// TIA Portal V20 export
VAR_GLOBAL   // PLC tag table "standard"
   SIMULACE AT %M2.0 : Bool;
   LOG_0 AT %M2.1 : Bool;
   LOG_1 AT %M2.2 : Bool;
   SMAZ_ME_0 AT %M2.3 : Bool;
   SMAZ_ME_1 AT %M2.4 : Bool;
   AUTOMAT AT %M2.5 : Bool;
   MANUAL AT %M2.6 : Bool;
   INICIALIZACE_OK AT %M3.3 : Bool;
   INICIALIZACE AT %M3.4 : Bool;
   INICIALIZACE_RUN AT %M3.5 : Bool;
   LINE_READY_START AT %M3.6 : Bool;
   alrm_global AT %M3.2 : Bool;
   wrong_global AT %M3.7 : Bool;
   alrm_op_0 AT %M4.0 : Bool;
   wrong_op_0 AT %M4.1 : Bool;
   alrm_op_1 AT %M4.2 : Bool;
   wrong_op_1 AT %M4.3 : Bool;
   I_i AT %MW6 : Int;
   "I_i(1)" AT %MW8 : Int;
   adresace AT %MW12 : Int;
   byte_smazat AT %MB5 : Byte;
   inicializace_block AT %M4.4 : Bool;
   s2_hsc_hrana AT %M4.5 : Bool;
   hodnota_volitelna AT %MB14 : Byte;
   Clock_Byte AT %MB0 : Byte;
   Clock_10Hz AT %M0.0 : Bool;
   Clock_5Hz AT %M0.1 : Bool;
   "Clock_2.5Hz" AT %M0.2 : Bool;
   Clock_2Hz AT %M0.3 : Bool;
   "Clock_1.25Hz" AT %M0.4 : Bool;
   Clock_1Hz AT %M0.5 : Bool;
   "Clock_0.625Hz" AT %M0.6 : Bool;
   "Clock_0.5Hz" AT %M0.7 : Bool;
   System_Byte AT %MB1 : Byte;
   FirstScan AT %M1.0 : Bool;
   DiagStatusUpdate AT %M1.1 : Bool;
   AlwaysTRUE AT %M1.2 : Bool;
   AlwaysFALSE AT %M1.3 : Bool;
   INICIALIZACE_REPEAT AT %M4.6 : Bool;
   AUT_MAN_HMI AT %M4.7 : Bool;   // POUŽÍVÁNO PRO PANELOUVOU VOLBU
   volny_pristup_2 AT %M10.0 : Bool;
   alrm_op_2 AT %M11.3 : Bool;
   wrong_op_2 AT %M11.4 : Bool;
   alrm_op_3 AT %M11.5 : Bool;
   wrong_op_3 AT %M11.6 : Bool;
   alrm_op_4 AT %M11.7 : Bool;
   wrong_op_4 AT %M15.0 : Bool;
   alrm_op_5 AT %M15.1 : Bool;
   wrong_op_5 AT %M15.2 : Bool;
   citac AT %M15.4 : Bool;
END_VAR
